(* PLC project types, tcpethernet types 1 *)
(* stored: creationDateTime 2026-10-28T09:00:00, modificationDateTime 2026-10-28T09:00:00 *)

TYPE Point : STRUCT
  x : INT := 1;
  y : INT;
END_STRUCT;
END_TYPE

TYPE Mode : (Idle, Running := 5);
END_TYPE

TYPE Buffer : ARRAY[0..3] OF INT := [10, 3(2)];
END_TYPE

TYPE Speed : INT := 7;
END_TYPE

FUNCTION Twice : INT
  VAR_INPUT
    v : INT;
  END_VAR

            Twice := v * 2;
          
END_FUNCTION

PROGRAM main
  VAR
    p : Point := (y := 4);
    m : Mode;
    buf : Buffer;
    s : Speed;
    sum : INT;
    scans : DINT;
  END_VAR

            scans := scans + 1;
IF scans > 1 THEN
  m := Mode#Running;
END_IF;
sum := Twice(p.x + p.y) + buf[0] + buf[3] + s;
          
END_PROGRAM
